(* CODESYS project textmaster.library
   Company: KOSTAL GmbH & Co.KG
   DefaultNamespace: KOSTAL.AF2024.Templates.TextMaster
   Version: 1.0.0.0
   Placeholder: KOSTAL.AF2024.Templates.TextMaster
   Author: M. Hundt
   Title: KOSTAL.AF2024.Templates.TextMaster

Project tree, tasks and I/O mapping:
  libraries: KOSTAL.AF2024.Core.FileLogger, 1.0.0.0 (KOSTAL GmbH & Co.KG); KOSTAL.AF2024.Core.ID, 1.0.0.0 (KOSTAL GmbH & Co.KG); KOSTAL.AF2024.Core.MainControl, 1.0.0.0 (KOSTAL GmbH & Co.KG); KOSTAL.AF2024.Core.Process, 1.0.0.0 (KOSTAL GmbH & Co.KG); KOSTAL.AF2024.Core.Settings, 1.0.0.0 (KOSTAL GmbH & Co.KG); KOSTAL.AF2024.Core.Station, 1.0.0.0 (KOSTAL GmbH & Co.KG); KOSTAL.AF2024.Core.StringTools, 1.0.0.0 (KOSTAL GmbH & Co.KG); KOSTAL.AF2024.Core.Text, 1.0.0.0 (KOSTAL GmbH & Co.KG); KOSTAL.AF2024.HMI.Controls, 1.0.0.0 (KOSTAL GmbH & Co.KG); KOSTAL.AF2024.HMI.I_Hmi, 1.0.0.0 (KOSTAL GmbH & Co.KG); Tc2_Standard, 3.3.3.0 (Beckhoff Automation GmbH)
  function block FB_TextMaster [ST]: _HmiDefine, _log_Start, _logLanguage, _mText, _mTextCommon, _parameterControl, _resetCondition, _getNameAndID, _ID_TO_WSTRING, _log, Condition, Condition_Owner, FB_init, ID, LogText, Message, Message_Owner, Name, TextPath, _linkHmi, FBmain, MasterPath, Path, SelectedLanguage, Text
  function block T_E_Text_TextMaster [ST]: Execution, failed, inProcess, Language, Name, notAccepted, NoTextLoaded, ReadText_0, Restart, TextAvailable
*)

// FB_TextMaster
FUNCTION_BLOCK Abstract FB_TextMaster IMPLEMENTS KOSTAL_AF2024_Core_Station.I_Station_Free, KOSTAL_AF2024_Core_Station.I_Station_Free_Owner //EXTENDS KOSTAL_AF2024_Core_Station.FB_Station_Free


VAR
	//From Station
	//=============================================================================================================================================================
	_ID	: KOSTAL_AF2024_Core_ID.T_ID;

	_Name	: KOSTAL_AF2024_Core_Settings.T_MaxString;	//localized name of station

	_condition			: KOSTAL_AF2024_Core_Process.FB_processCondition;

	_Logger	: KOSTAL_AF2024_Core_FileLogger.I_Logger;
	
	_message				: KOSTAL_AF2024_Core_Process.T_messageText_3_lines;
	//=============================================================================================================================================================

	//TextMaster	
	//=============================================================================================================================================================

	_pathCommon	: KOSTAL_AF2024_Core_Settings.T_MaxString_UTF8;
	
	
	//"Master" Text provider with Common content for the whole project
	_TextCommon	: KOSTAL_AF2024_Core_Text.FB_Handler_Master;

//	//"Slave" local text provider for FB_TextMaster only
	_TextPath		: KOSTAL_AF2024_Core_Settings.T_MaxString_UTF8;
	_Text	: KOSTAL_AF2024_Core_Text.FB_Handler_Slave;
	
	_E_Text		: T_E_Text_TextMaster;
	
	_iHmi_station				: KOSTAL_AF2024_HMI_I_Hmi.I_Page_Station_Owner; //KOSTAL_AF2024_HMI_WinHMI.FB_Page_Station;	 

	_loggedText: KOSTAL_AF2024_Core_Settings.T_MaxString;

	_logStart	: BOOL:= TRUE;
	//=============================================================================================================================================================

END_VAR

METHOD PROTECTED _HmiDefine
VAR_INPUT
END_VAR
//_HMI_station.FBmain();


_Name:= _Text.GetText(_E_Text.Name);


_iHmi_station.Name:= _Name;
     
_iHmi_station.Text.line_01:= _condition.message.line_01;
_iHmi_station.Text.line_02:= _condition.message.line_02;
_iHmi_station.Text.line_03:= _condition.message.line_03;
     
_iHmi_station.Button_Escape.Visible	:= _condition.isError() OR _iHmi_station.Button_Escape.Sign;
_iHmi_station.Button_Escape.Text		:= _Text.GetText(_E_Text.Restart);
     
_iHmi_station.Status.CopyFrom(_condition);
END_METHOD

METHOD PROTECTED _log_Start : BOOL
VAR_INPUT
END_VAR

IF _logStart AND _Text.State.ready AND (_Text.LoadedLanguage <> '') THEN

	IF _log("===START===") THEN	_LogStart:= FALSE;	END_IF

END_IF
END_METHOD

METHOD PROTECTED _logLanguage
VAR_INPUT
END_VAR

IF _TextCommon.LoadedLanguage = ''										
	THEN RETURN;	
END_IF
IF _TextCommon.LoadedLanguage <> _Text.LoadedLanguage	
	THEN RETURN;	
END_IF
IF _loggedText = STRING_TO_WSTRING(_Text.LoadedLanguage)						THEN RETURN;	END_IF

IF _log(STRING_TO_WSTRING(TC2_Standard.CONCAT('Language changed to ', _TextCommon.LoadedLanguage)))	THEN
	_loggedText:= STRING_TO_WSTRING(_TextCommon.LoadedLanguage);
END_IF
END_METHOD

//local text
METHOD PROTECTED _mText
VAR_INPUT
END_VAR

_Text.Path:= _textPath;// Tc2_Standard.CONCAT(GVL_FilesAndFolder.PROJEKT_PATH, _PATH_SLAVE);
_Text.FBmain();
END_METHOD

METHOD PROTECTED _mTextCommon

_TextCommon.Path:= _pathCommon;// Tc2_Standard.CONCAT(GVL_FilesAndFolder.PROJEKT_PATH, _PATH_MASTER);
_TextCommon.FBmain();
END_METHOD

METHOD PROTECTED _parameterControl : BOOL
VAR_INPUT
END_VAR

_parameterControl:= FALSE;

IF _iHmi_station = 0 THEN

	_message.clear();
	_message.line_01:= "Link missing";
	_message.line_02:= "Interface _iHmi is not linked";

	_condition.setMessage(4999, _message);

ELSE

	_parameterControl:= TRUE;

END_IF
END_METHOD

METHOD PROTECTED _resetCondition
VAR_INPUT
END_VAR

IF _condition.isText() THEN
	_condition.clear();
ELSIF _condition.isInfo() THEN
	_condition.clear();
ELSIF _condition.isMessage() THEN
	_condition.clear();
ELSIF _condition.isMasterMessage() THEN
	_condition.clear();
ELSIF _iHmi_station.Button_Escape.Pulse THEN
	_log(_condition.Message.toString());
	_condition.clear();
END_IF
END_METHOD

METHOD PROTECTED _getNameAndID : KOSTAL_AF2024_Core_Settings.T_MaxString

VAR
	_c	: KOSTAL_AF2024_Core_StringTools.FB_Concat;
END_VAR


_c.Clear();
_c.addContent(_Name);
_c.addContent("[");
_c.addContent(_ID.name);
_c.addContent("(");
_c.addContent(DINT_TO_WSTRING(_ID.key));
_c.addContent(")");
_c.addContent("]");
_getNameAndID:= _c.getResult();
_c.Clear();
END_METHOD

METHOD PROTECTED _ID_TO_WSTRING : KOSTAL_AF2024_Core_Settings.T_MaxString

VAR
	_c	: KOSTAL_AF2024_Core_StringTools.FB_Concat;
END_VAR


_c.Clear();
_c.addContent(_ID.name);
_c.addContent("(");
_c.addContent(DINT_TO_WSTRING(_ID.key));
_c.addContent(")");
_ID_TO_WSTRING:= _c.getResult();
_c.Clear();
END_METHOD

METHOD PROTECTED _log : BOOL
VAR_INPUT
	Text	: KOSTAL_AF2024_Core_Settings.T_MaxString;
END_VAR

IF _Logger = 0 THEN 
	RETURN;	
END_IF
IF NOT _Logger.State.success THEN 
	RETURN;	
END_IF

_Logger.ID					:= _ID_TO_WSTRING();
_Logger.name				:= _Name;


_Logger.addLine(Text);

_log:= TRUE;
END_METHOD

PROPERTY PUBLIC Condition : KOSTAL_AF2024_Core_Process.I_processCondition
GET

Condition := _condition;
END_GET
END_PROPERTY

PROPERTY PUBLIC Condition_Owner : KOSTAL_AF2024_Core_Process.I_processCondition_Owner
GET

Condition_Owner := _condition;
END_GET
END_PROPERTY

METHOD FB_init : BOOL
VAR_INPUT
	bInitRetains 	: BOOL; // if TRUE, the retain variables are initialized (warm start / cold start)
	bInCopyCode 	: BOOL;  // if TRUE, the instance afterwards gets moved into the copy code (online change)
	ID_Name				: KOSTAL_AF2024_Core_Settings.T_MaxString;
	ID_Key				: DINT;
END_VAR

_ID.name:= ID_Name;
_ID.key	:= ID_Key;
END_METHOD

PROPERTY PUBLIC ID : KOSTAL_AF2024_Core_ID.I_T_ID
GET

ID := _ID;
END_GET
END_PROPERTY

(*
	These PUBLIC methods are required to make the log function usable for interface participants (such as cylinders).
*)
METHOD PUBLIC LogText : BOOL
VAR_INPUT
	Text	: KOSTAL_AF2024_Core_Settings.T_MaxString;
END_VAR
LogText:= _log(Text);
END_METHOD

PROPERTY PUBLIC Message : KOSTAL_AF2024_Core_Process.I_T_messageText_3_lines
GET

Message := _message;
END_GET
END_PROPERTY

PROPERTY PUBLIC Message_Owner : KOSTAL_AF2024_Core_Process.I_T_messageText_3_lines_Owner
GET

Message_Owner := _message;
END_GET
END_PROPERTY

//localized name of station
PROPERTY PUBLIC Name : KOSTAL_AF2024_Core_Settings.T_MaxString
GET

Name:= _Name;
END_GET
SET

_Name:= Name;
END_SET
END_PROPERTY

PROPERTY PUBLIC TextPath : KOSTAL_AF2024_Core_Settings.T_MaxString_UTF8
GET

TextPath:= _TextPath;
END_GET
SET

_TextPath:= TextPath;
END_SET
END_PROPERTY

METHOD PROTECTED ABSTRACT _linkHmi
VAR_INPUT
END_VAR
END_METHOD

METHOD PUBLIC FBmain


VAR
	_udi: UDINT;
END_VAR
_linkHmi();

IF NOT _parameterControl()	THEN RETURN;	END_IF

_HmiDefine();

_resetCondition();

_mTextCommon();

_mText();

_log_Start();

_logLanguage();

IF _pathCommon = '' THEN
	_message.clear();
	_message.line_01	:=	"Text loading failed";
	_message.line_02	:=	"Common path Missing";
	_condition.setMessage(KOSTAL_AF2024_Core_process.E_PROCESS_CONDITION_DEFAULT_PRIORITYLEVEL.ERROR, _message);
	
ELSIF _TextPath = '' THEN
	_message.clear();
	_message.line_01	:=	"Text loading failed";
	_message.line_02	:=	"Text path Missing";
	_condition.setMessage(KOSTAL_AF2024_Core_process.E_PROCESS_CONDITION_DEFAULT_PRIORITYLEVEL.ERROR, _message);
ELSIF _TextCommon.State.fail THEN

	_message.clear();

	IF _Text.State.ready AND (_Text.LoadedLanguage <> '')	THEN	

		_Text.ClearVars();
		_Text.AddVar(_Text.GetText(_E_Text.failed));
		_message.line_01	:=	_Text.GetText(_E_Text.ReadText_0);

	ELSE	
		_message.line_01	:=	"Text loading failed";
	END_IF
	
	_message.line_02	:=	_TextCommon.State.description;

	IF NOT _condition.isError() THEN _log(_Message.toString());	END_IF
	_condition.setMessage(KOSTAL_AF2024_Core_process.E_PROCESS_CONDITION_DEFAULT_PRIORITYLEVEL.ERROR, _message);

ELSIF NOT _TextCommon.State.ready THEN

	_message.clear();
	
	IF _Text.State.ready AND (_Text.LoadedLanguage <> '')	THEN	

		_Text.ClearVars();
		_Text.AddVar(_Text.GetText(_E_Text.inProcess));
		_message.line_01	:=	_Text.GetText(_E_Text.ReadText_0);
			
	ELSE	_message.line_01			:=	"Text loading in process";
	END_IF

	_message.line_02	:=	_TextCommon.State.description;

	_condition.setMessage(KOSTAL_AF2024_Core_process.E_PROCESS_CONDITION_DEFAULT_PRIORITYLEVEL.MESSAGE, _message);

ELSIF _TextCommon.LoadedLanguage = '' THEN

	_message.clear();

	IF _Text.State.ready AND (_Text.LoadedLanguage <> '')	THEN	
		_message.line_01	:=	_Text.GetText(_E_Text.NoTextLoaded);
	ELSE
		_message.line_01	:=	"No Text available";
	END_IF

	_message.line_02	:=	_TextCommon.State.description;

	_condition.setMessage(KOSTAL_AF2024_Core_process.E_PROCESS_CONDITION_DEFAULT_PRIORITYLEVEL.MESSAGE, _message);

	
ELSE
	
	_message.clear();
	IF _Text.State.ready AND (_Text.LoadedLanguage <> '')	THEN	_message.line_01	:=	_Text.GetText (_E_Text.TextAvailable);
	ELSE																													_message.line_01	:=	"Text available";
	END_IF
	
	_message.line_02	:=	_TextCommon.State.description;

	_condition.setMessage(KOSTAL_AF2024_Core_process.E_PROCESS_CONDITION_DEFAULT_PRIORITYLEVEL.INFORMATION, _message);

END_IF
END_METHOD

PROPERTY PUBLIC MasterPath : KOSTAL_AF2024_Core_Settings.T_MaxString_UTF8
GET
MasterPath := _pathCommon;
END_GET
SET
_pathCommon := MasterPath;
END_SET
END_PROPERTY

PROPERTY PUBLIC Path : KOSTAL_AF2024_Core_Settings.T_MaxString_UTF8
GET

Path:= _TextCommon.Path;
END_GET
END_PROPERTY

PROPERTY PUBLIC SelectedLanguage : KOSTAL_AF2024_Core_Settings.T_MaxString_UTF8
GET

SelectedLanguage:= _TextCommon.SelectedLanguage;
END_GET
SET

_TextCommon.SelectedLanguage:= SelectedLanguage;
END_SET
END_PROPERTY

PROPERTY PUBLIC Text : KOSTAL_AF2024_Core_Text.I_Text
GET

Text:= _TextCommon;
END_GET
END_PROPERTY

END_FUNCTION_BLOCK

// T_E_Text_TextMaster
FUNCTION_BLOCK T_E_Text_TextMaster EXTENDS KOSTAL_AF2024_Core_Text.T_E_Text
VAR_INPUT
END_VAR
VAR_OUTPUT
END_VAR
VAR
END_VAR

PROPERTY Execution : ST_E_Text
GET

Execution.Number:= 8;
END_GET
END_PROPERTY

PROPERTY failed : ST_E_Text
GET

failed.Number:= 7;
END_GET
END_PROPERTY

PROPERTY inProcess : ST_E_Text
GET

inProcess.Number:= 6;
END_GET
END_PROPERTY

PROPERTY Language : ST_E_Text
GET

Language.Number:= 1;
END_GET
END_PROPERTY

PROPERTY Name : ST_E_Text
GET

Name.Number:= 2;
END_GET
END_PROPERTY

PROPERTY notAccepted : ST_E_Text
GET

notAccepted.Number:= 5;
END_GET
END_PROPERTY

PROPERTY NoTextLoaded : ST_E_Text
GET

NoTextLoaded.Number:= 9;
END_GET
END_PROPERTY

PROPERTY ReadText_0 : ST_E_Text
GET

ReadText_0.Number:= 4;
END_GET
END_PROPERTY

PROPERTY Restart : ST_E_Text
GET

Restart.Number:= 3;
END_GET
END_PROPERTY

PROPERTY TextAvailable : ST_E_Text
GET

TextAvailable.Number:= 10;
END_GET
END_PROPERTY

END_FUNCTION_BLOCK
